RoboDK station: Rubiks_Meca500.rdk

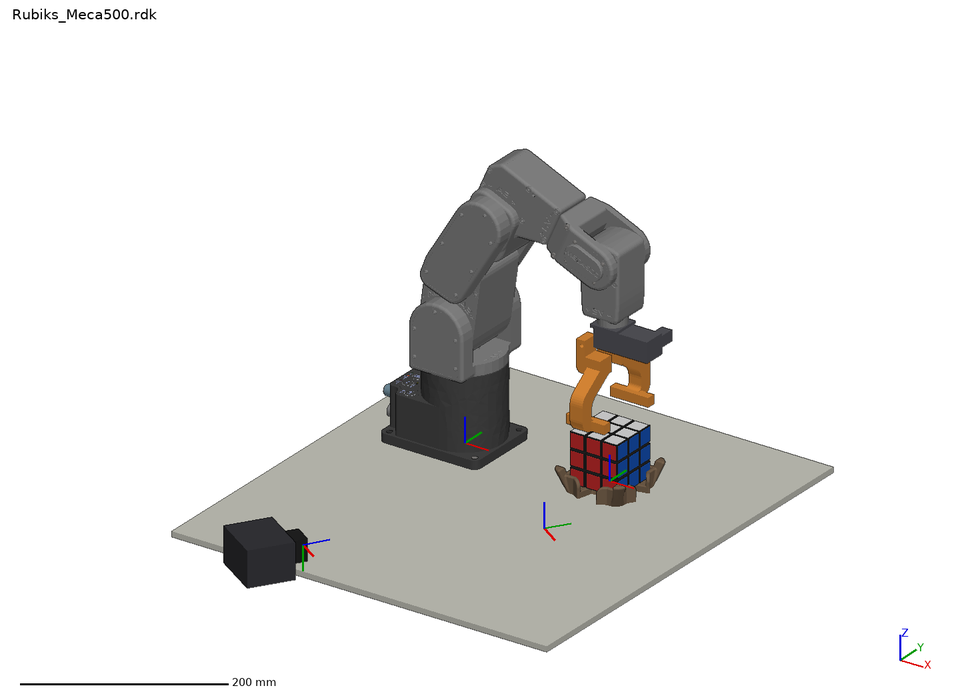
[picture v0: the station drawn from its stored meshes, robots at their saved joint values, targets as dots, program paths as lines]
Station Rubiks Meca500 (saved by RoboDK 6.0.7). Poses are relative to the parent item; angles as X-Y-Z fixed-axis rotations.
  - frame Mecademic Meca500 R3 Base at (0, 0, 0) mm
    - robot Mecademic Meca500 R3: 6 axes
        modified DH rows (alpha deg, a mm, theta deg, d mm): 0, 0, 0, 135; -90, 0, -90, 0; 0, 135, 0, 0; -90, 38, 0, 120; 90, 0, 0, 0; -90, 0, 180, 70
        joint limits [-175, -70, -135, -170, -115, -720] to [175, 90, 70, 170, 115, 720]; home [0, 0, 0, 0, 0, 0]; saved at [0, 20.83, 3.116, 0, 66.054, 0]
      - tool MEGP 25E, TCP at (3.1, 0, 93.2) mm
        - object Pince at (-3.1, 0, -93.2) mm, size 70 x 45.2 x 25.4 mm
        - object Doigt_1 at (-22.47, 56.8, 5.03) mm, rotated rx -90 ry 0 rz -90 deg, size 48.3 x 85.2 x 45 mm, geometry from mors.STL
        - object Doigt_2 at (-22.47, 34.8, 5.03) mm, rotated rx -90 ry 0 rz -90 deg, size 48.3 x 85.2 x 45 mm, geometry from Mors_droite.STL
    - frame Socle_repere at (170, 0, 7) mm
      - object Socle at (0, 0, 0) mm, size 81.4 x 81.4 x 25.5 mm, geometry from socle.stl
      - object Cubie_-1-1-1 at (-19, -19, 9.5) mm, size 17.9 x 17.9 x 17.9 mm
      - object Cubie_-1-1+0 at (-19, -19, 28.5) mm, size 17.9 x 17.9 x 17.4 mm
      - object Cubie_-1-1+1 at (-19, -19, 47.5) mm, size 17.9 x 17.9 x 17.9 mm
      - object Cubie_-1+0-1 at (-19, 0, 9.5) mm, size 17.9 x 17.4 x 17.9 mm
      - object Cubie_-1+0+0 at (-19, 0, 28.5) mm, size 17.9 x 17.4 x 17.4 mm
      - object Cubie_-1+0+1 at (-19, 0, 47.5) mm, size 17.9 x 17.4 x 17.9 mm
      - object Cubie_-1+1-1 at (-19, 19, 9.5) mm, size 17.9 x 17.9 x 17.9 mm
      - object Cubie_-1+1+0 at (-19, 19, 28.5) mm, size 17.9 x 17.9 x 17.4 mm
      - object Cubie_-1+1+1 at (-19, 19, 47.5) mm, size 17.9 x 17.9 x 17.9 mm
      - object Cubie_+0-1-1 at (0, -19, 9.5) mm, size 17.4 x 17.9 x 17.9 mm
      - object Cubie_+0-1+0 at (0, -19, 28.5) mm, size 17.4 x 17.9 x 17.4 mm
      - object Cubie_+0-1+1 at (0, -19, 47.5) mm, size 17.4 x 17.9 x 17.9 mm
      - object Cubie_+0+0-1 at (0, 0, 9.5) mm, size 17.4 x 17.4 x 17.9 mm
      - object Cubie_+0+0+1 at (0, 0, 47.5) mm, size 17.4 x 17.4 x 17.9 mm
      - object Cubie_+0+1-1 at (0, 19, 9.5) mm, size 17.4 x 17.9 x 17.9 mm
      - object Cubie_+0+1+0 at (0, 19, 28.5) mm, size 17.4 x 17.9 x 17.4 mm
      - object Cubie_+0+1+1 at (0, 19, 47.5) mm, size 17.4 x 17.9 x 17.9 mm
      - object Cubie_+1-1-1 at (19, -19, 9.5) mm, size 17.9 x 17.9 x 17.9 mm
      - object Cubie_+1-1+0 at (19, -19, 28.5) mm, size 17.9 x 17.9 x 17.4 mm
      - object Cubie_+1-1+1 at (19, -19, 47.5) mm, size 17.9 x 17.9 x 17.9 mm
      - object Cubie_+1+0-1 at (19, 0, 9.5) mm, size 17.9 x 17.4 x 17.9 mm
      - object Cubie_+1+0+0 at (19, 0, 28.5) mm, size 17.9 x 17.4 x 17.4 mm
      - object Cubie_+1+0+1 at (19, 0, 47.5) mm, size 17.9 x 17.4 x 17.9 mm
      - object Cubie_+1+1-1 at (19, 19, 9.5) mm, size 17.9 x 17.9 x 17.9 mm
      - object Cubie_+1+1+0 at (19, 19, 28.5) mm, size 17.9 x 17.9 x 17.4 mm
      - object Cubie_+1+1+1 at (19, 19, 47.5) mm, size 17.9 x 17.9 x 17.9 mm
    - frame Table_repere at (170, -110, 0) mm, rotated rx 0 ry 0 rz -32.91 deg
      - frame Camera_repere at (0, -250, 28.5) mm, rotated rx -90 ry 0 rz 0 deg
        - object Camera at (0, 0, 0) mm, size 60 x 48.5 x 70 mm
    - object Table at (0, 0, 0) mm, size 440 x 480 x 6 mm
  - Python program remise_a_zero (listed below)
  - Python program verifier_mouvements (listed below)
  - Python program verifier_outil (listed below)
  - Python program prendre_et_reposer (listed below)
  - Python program tourner_cube_gauche (listed below)
  - Python program tourner_cube_droite (listed below)
  - Python program basculer_gauche (listed below)
  - Python program basculer_droite (listed below)
  - Python program basculer_avant (listed below)
  - Python program basculer_arriere (listed below)
  - Python program tourner_haut_gauche (listed below)
  - Python program tourner_haut_droite (listed below)
  - Python program tourner_haut_demi_tour (listed below)
  - Python program presenter_faces (listed below)

--- Python program remise_a_zero ---
# -*- coding: utf-8 -*-
# Programme RoboDK : exécute meca500_rubiks.remise_a_zero() dans la simulation.
import os
import sys
from robodk import robolink
projet = robolink.Robolink().getParam("PATH_OPENSTATION")    # dossier de Rubiks_Meca500.rdk
sys.path.insert(0, os.path.join(projet, "simulation"))
import simulateur
simulateur.simuler('remise_a_zero')

--- Python program verifier_mouvements ---
# -*- coding: utf-8 -*-
# Programme RoboDK : exécute meca500_rubiks.verifier_mouvements() dans la simulation.
import os
import sys
from robodk import robolink
projet = robolink.Robolink().getParam("PATH_OPENSTATION")    # dossier de Rubiks_Meca500.rdk
sys.path.insert(0, os.path.join(projet, "simulation"))
import simulateur
simulateur.simuler('verifier_mouvements')

--- Python program verifier_outil ---
# -*- coding: utf-8 -*-
# Programme RoboDK : exécute meca500_rubiks.verifier_outil() dans la simulation.
import os
import sys
from robodk import robolink
projet = robolink.Robolink().getParam("PATH_OPENSTATION")    # dossier de Rubiks_Meca500.rdk
sys.path.insert(0, os.path.join(projet, "simulation"))
import simulateur
simulateur.simuler('verifier_outil')

--- Python program prendre_et_reposer ---
# -*- coding: utf-8 -*-
# Programme RoboDK : exécute meca500_rubiks.prendre_et_reposer() dans la simulation.
import os
import sys
from robodk import robolink
projet = robolink.Robolink().getParam("PATH_OPENSTATION")    # dossier de Rubiks_Meca500.rdk
sys.path.insert(0, os.path.join(projet, "simulation"))
import simulateur
simulateur.simuler('prendre_et_reposer')

--- Python program tourner_cube_gauche ---
# -*- coding: utf-8 -*-
# Programme RoboDK : exécute meca500_rubiks.tourner_cube_gauche() dans la simulation.
import os
import sys
from robodk import robolink
projet = robolink.Robolink().getParam("PATH_OPENSTATION")    # dossier de Rubiks_Meca500.rdk
sys.path.insert(0, os.path.join(projet, "simulation"))
import simulateur
simulateur.simuler('tourner_cube_gauche')

--- Python program tourner_cube_droite ---
# -*- coding: utf-8 -*-
# Programme RoboDK : exécute meca500_rubiks.tourner_cube_droite() dans la simulation.
import os
import sys
from robodk import robolink
projet = robolink.Robolink().getParam("PATH_OPENSTATION")    # dossier de Rubiks_Meca500.rdk
sys.path.insert(0, os.path.join(projet, "simulation"))
import simulateur
simulateur.simuler('tourner_cube_droite')

--- Python program basculer_gauche ---
# -*- coding: utf-8 -*-
# Programme RoboDK : exécute meca500_rubiks.basculer_gauche() dans la simulation.
import os
import sys
from robodk import robolink
projet = robolink.Robolink().getParam("PATH_OPENSTATION")    # dossier de Rubiks_Meca500.rdk
sys.path.insert(0, os.path.join(projet, "simulation"))
import simulateur
simulateur.simuler('basculer_gauche')

--- Python program basculer_droite ---
# -*- coding: utf-8 -*-
# Programme RoboDK : exécute meca500_rubiks.basculer_droite() dans la simulation.
import os
import sys
from robodk import robolink
projet = robolink.Robolink().getParam("PATH_OPENSTATION")    # dossier de Rubiks_Meca500.rdk
sys.path.insert(0, os.path.join(projet, "simulation"))
import simulateur
simulateur.simuler('basculer_droite')

--- Python program basculer_avant ---
# -*- coding: utf-8 -*-
# Programme RoboDK : exécute meca500_rubiks.basculer_avant() dans la simulation.
import os
import sys
from robodk import robolink
projet = robolink.Robolink().getParam("PATH_OPENSTATION")    # dossier de Rubiks_Meca500.rdk
sys.path.insert(0, os.path.join(projet, "simulation"))
import simulateur
simulateur.simuler('basculer_avant')

--- Python program basculer_arriere ---
# -*- coding: utf-8 -*-
# Programme RoboDK : exécute meca500_rubiks.basculer_arriere() dans la simulation.
import os
import sys
from robodk import robolink
projet = robolink.Robolink().getParam("PATH_OPENSTATION")    # dossier de Rubiks_Meca500.rdk
sys.path.insert(0, os.path.join(projet, "simulation"))
import simulateur
simulateur.simuler('basculer_arriere')

--- Python program tourner_haut_gauche ---
# -*- coding: utf-8 -*-
# Programme RoboDK : exécute meca500_rubiks.tourner_haut_gauche() dans la simulation.
import os
import sys
from robodk import robolink
projet = robolink.Robolink().getParam("PATH_OPENSTATION")    # dossier de Rubiks_Meca500.rdk
sys.path.insert(0, os.path.join(projet, "simulation"))
import simulateur
simulateur.simuler('tourner_haut_gauche')

--- Python program tourner_haut_droite ---
# -*- coding: utf-8 -*-
# Programme RoboDK : exécute meca500_rubiks.tourner_haut_droite() dans la simulation.
import os
import sys
from robodk import robolink
projet = robolink.Robolink().getParam("PATH_OPENSTATION")    # dossier de Rubiks_Meca500.rdk
sys.path.insert(0, os.path.join(projet, "simulation"))
import simulateur
simulateur.simuler('tourner_haut_droite')

--- Python program tourner_haut_demi_tour ---
# -*- coding: utf-8 -*-
# Programme RoboDK : exécute meca500_rubiks.tourner_haut_demi_tour() dans la simulation.
import os
import sys
from robodk import robolink
projet = robolink.Robolink().getParam("PATH_OPENSTATION")    # dossier de Rubiks_Meca500.rdk
sys.path.insert(0, os.path.join(projet, "simulation"))
import simulateur
simulateur.simuler('tourner_haut_demi_tour')

--- Python program presenter_faces ---
# -*- coding: utf-8 -*-
# Programme RoboDK : exécute meca500_rubiks.presenter_faces() dans la simulation.
import os
import sys
from robodk import robolink
projet = robolink.Robolink().getParam("PATH_OPENSTATION")    # dossier de Rubiks_Meca500.rdk
sys.path.insert(0, os.path.join(projet, "simulation"))
import simulateur
simulateur.simuler('presenter_faces')
